TYPE ST_ActuatorModulatingFunctions :
STRUCT
	ToPosition			: FB_SequencerFunction; //param E_ActuatorModulatingFunctionParam.Position
	Open				: FB_SequencerFunction;
	Close				: FB_SequencerFunction;
END_STRUCT
END_TYPE

(* stored: Version 1.1.0.1, ProductVersion 3.1.4024.12
   DUT ST_ActuatorModulatingFunctions: Id {abc305ee-6736-445a-8d8d-6f85cdc8a017} *)
